// TwinCAT 3 PLC project Untitled1
// ProgramVersion: 3.1.4024.0
// libraries:
//   Tc2_Standard, * (Beckhoff Automation GmbH)
//   Tc2_System, * (Beckhoff Automation GmbH)
//   Tc3_Module, * (Beckhoff Automation GmbH)
// project tree:
//   / GlobalTextList.TcGTLO, PlcTask.TcTTO, Visualization Manager.TcVMO (not stored)
//   GVLs/ GVL_IO.TcGVL, GVL_SAFETY.TcGVL
//   POUs/ MAIN.TcPOU
//   VISUs/ Visualization.TcVIS
// real-time tasks:
//   TASK PlcTask: cycle T#10ms, priority 20, ADS port 350
// I/O:
//   DEVICE Device 1 (EtherCAT), AmsNetId 5.34.198.36.2.1
//     Term 1 (EK1200) [EK1200-5000 EtherCAT Power supply (2A E-Bus)]
//       Term 2 (EL6910) [EL6910, TwinSAFE PLC]
//       Term 3 (EL1904) [EL1904, 4 Ch. Safety Input 24V, TwinSAFE]
//         modules: Module 1 (FSOES)
//       Term 4 (EL9011) [EL9011 End Terminal]
//   DEVICE Device 5 (EtherCAT), AmsNetId 5.34.198.36.6.1
//     Box 5 (KRC4 secondary EL6695-1001) [KRC4 secondary EL6695-1001]
//       modules: Module 1 (Sync Inputs), Module 2 (Safety Data Bitf  (8 Byte)), Module 3 (Default IO)
// variable links:
//   Device 1 (EtherCAT) <-> Device 5 (EtherCAT)/Box 5 (KRC4 secondary EL6695-1001)
//     Term 1 (EK1200)/Term 2 (EL6910)/ConnectionInputs/Message_5 TxPDO <-> Module 2 (Safety Data Bitf  (8 Byte))/Outputs Bitf/FSOE
//   Device 5 (EtherCAT) <-> Device 1 (EtherCAT)/Term 1 (EK1200)/Term 2 (EL6910)
//     Box 5 (KRC4 secondary EL6695-1001)/Module 2 (Safety Data Bitf  (8 Byte))/Inputs Bitf/FSOE <-> ConnectionOutputs/Message_5 RxPDO
//   (this object) <-> Device 1 (EtherCAT)
//     Term 1 (EK1200)/Term 2 (EL6910)/ConnectionInputs/Message_3 TxPDO <-> Term 1 (EK1200)/Term 3 (EL1904)/Module 1 (FSOES)/RxPDO/FSOE
//     Term 1 (EK1200)/Term 2 (EL6910)/ConnectionOutputs/Message_3 RxPDO <-> Term 1 (EK1200)/Term 3 (EL1904)/Module 1 (FSOES)/TxPDO/FSOE
//     Term 1 (EK1200)/Term 3 (EL1904)/Module 1 (FSOES)/RxPDO/FSOE <-> Term 1 (EK1200)/Term 2 (EL6910)/ConnectionInputs/Message_3 TxPDO
//     Term 1 (EK1200)/Term 3 (EL1904)/Module 1 (FSOES)/TxPDO/FSOE <-> Term 1 (EK1200)/Term 2 (EL6910)/ConnectionOutputs/Message_3 RxPDO
//   Untitled1 Instance <-> Device 1 (EtherCAT)/Term 1 (EK1200)/Term 2 (EL6910)
//     PlcTask Inputs/GVL_SAFETY.Estop1_Y <-> StandardInputs/Standard Out Var 4
//     PlcTask Inputs/GVL_SAFETY.bLocalEstopFromKUKA <-> StandardInputs/Standard Out Var 6
//     PlcTask Outputs/GVL_SAFETY.Estop1_RX <-> StandardOutputs/Standard In Var 1
//     PlcTask Outputs/GVL_SAFETY.bRunStop <-> StandardOutputs/Standard In Var 2

CONFIGURATION Untitled1
    RESOURCE PLC ON TwinCAT3
        TASK PlcTask(INTERVAL := T#10ms, PRIORITY := 20);
        PROGRAM MAIN WITH PlcTask : MAIN;
    END_RESOURCE
END_CONFIGURATION

// ---- GVLs/GVL_IO.TcGVL
VAR_GLOBAL
	Estop1_A AT %I* : BOOL ; (* Emergency stop 1 A-circuit NC *)
	Estop1_B AT %I* : BOOL ; (* Emergency stop 1 B-circuit NC *)
END_VAR

// ---- GVLs/GVL_SAFETY.TcGVL
VAR_GLOBAL
	Estop1_Y 				AT %I* 	: BOOL ; (* Emergency stop 1 status NC *)
	Estop1_RX 				AT %Q* 	: BOOL ; (* Restart emergency stop NO *)
	
	bLocalEstopFromKUKA 	AT %I* 	: BOOL ;
	bRunStop 				AT %Q*  : BOOL ;
END_VAR

// ---- POUs/MAIN.TcPOU
PROGRAM MAIN
VAR
	bCount : BOOL;
	iCounter : INT;
END_VAR

IF bCount THEN
	iCounter := iCounter + 1;
	GVL_SAFETY.bRunStop := TRUE;
END_IF;

END_PROGRAM

// ---- GlobalTextList.TcGTLO
TEXTLIST GlobalTextList
  898 = 'External'
  119 = 'Pendant'
  834 = 'Reset'
  761 = 'Run/Stop'
END_TEXTLIST

// ---- VISUs/Visualization.TcVIS
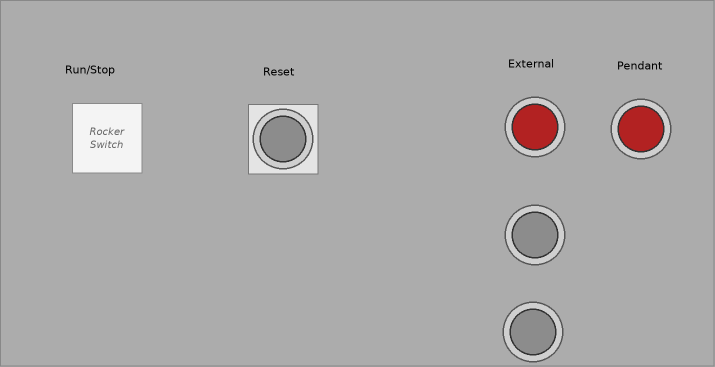
VISUALIZATION Visualization  // 715x367
    RockerSwitch (72,103 70x70), variable: bRunStop, behaviour: TOGGLE, style: Switch-RockerSwitch-Gray
    PushSwitch (248,104 70x70), variable: Estop1_RX, behaviour: TAP, style: Switch-PushSwitch-Gray
    Lamp1 (500,92 70x70), variable: not Estop1_Y, style: Lamp-Lamp1-Red
    Lamp1 (606,94 70x70), variable: not bLocalEstopFromKUKA, style: Lamp-Lamp1-Red
    Lamp1 (500,200 70x70), variable: Estop1_A, style: Lamp-Lamp1-Gray
    Lamp1 (498,297 70x70), variable: Estop1_B, style: Lamp-Lamp1-Gray
    Label (15,55 150x30), "Run/Stop"
    Label (204,57 150x30), "Reset"
    Label (456,49 150x30), "External"
    Label (565,51 150x30), "Pendant"
END_VISUALIZATION
